// TIA Portal project "Tables" (V21)

(* hardware
DEVICE "PLC_Tables"  S7-1500 station
   slot 0: "Rail_0"  Rack  6ES7 590-1***0-0AA0
   slot 1: "PLC_Tables"  CPU 1516-3 PN/DP  6ES7 516-3AN02-0AB0  V2.9
      slot 3: "CPU display_1"  6ES7591-1BA00-0AA0
      slot 32768: "PROFINET interface_1"  X1
         slot 32769: "Port_1"  X1 P1
         slot 32770: "Port_2"  X1 P2
      slot 33024: "PROFINET interface_2"  X2
         slot 33025: "Port_1"  X2 P1
      slot 33280: "DP interface_1"  X3
      slot 34817: "Virtual CP interface port_1"  Virtual CP interface port  Virtual CP interface port
*)

// ===== PLC "PLC_Tables"  CPU 1516-3 PN/DP =====
// protected blocks, not shown: "Sealed"

VAR_GLOBAL   // PLC tag table "IO"
   "Start" AT %I0.0 : Bool;   // Start button
   "Stop" AT %I0.1 : Bool;   // Stop button, normally closed
   "DoorClosed" AT %I0.2 : Bool;   // Door switch
   "Level" AT %IW2 : Int;   // Tank level in percent
   "Motor" AT %Q0.0 : Bool;   // Motor contactor
   "Lamp" AT %Q0.1 : Bool;   // Signal lamp
   "Valve" AT %Q0.2 : Bool;   // Inlet valve
   "Fault" AT %M0.0 : Bool;   // Collected fault
   "StartEdge" AT %M0.1 : Bool;   // Edge memory of Start
   "Setpoint" AT %MW10 : Int;   // Level setpoint
   "Parts" AT %MW12 : Int;   // Parts counted
   "Speed" AT %MD20 : Real;   // Conveyor speed
   "StatusWord" AT %MW30 : Word;   // Status bits
   "Alarm" AT %M1.0 : Bool;   // Set by the sealed block
END_VAR

TYPE "RecipeStep"
   STRUCT
      target : Real;   // Speed to reach
      duration : Time;   // How long to hold it
   END_STRUCT;
END_TYPE

// folder: Common

DATA_BLOCK "LampDelay"   // DB1
{ S7_Optimized_Access := 'TRUE' }
AUTHOR : Simatic
FAMILY : IEC
NAME : IEC_TMR
VERSION : 1.0
// stored: InstanceOfName IEC_TIMER
"IEC_TIMER"
BEGIN
END_DATA_BLOCK

// folder: Data

DATA_BLOCK "Recipe"   // DB2
{ S7_Optimized_Access := 'TRUE' }
VERSION : 0.1
   VAR
      active : Bool;   // A recipe runs
      count : Int;   // Cycles run
      steps : Array[1..3] of "RecipeStep";
      limits : Struct
         low : Int;
         high : Int := 90;
      END_STRUCT;
   END_VAR
BEGIN
END_DATA_BLOCK

DATA_BLOCK "LadBoxesData"   // DB3
{ S7_Optimized_Access := 'TRUE' }
VERSION : 0.1
// stored: InstanceOfName LadBoxes
"LadBoxes"
BEGIN
END_DATA_BLOCK

// folder: (top level)

ORGANIZATION_BLOCK "Main"   // OB1, SCL, ProgramCycle
TITLE = "Main Program Sweep (Cycle)"
{ S7_Optimized_Access := 'TRUE' }
VERSION : 0.1
   VAR_INPUT
      Initial_Call : Bool;   // Initial call of this OB
      Remanence : Bool;   // =True, if remanent data are available
   END_VAR
BEGIN

    "UseRecipe"();
    "Sealed"();
    "LadBoxesData"();
    "StatusWord" := "StatusWord" OR 16#0001;
END_ORGANIZATION_BLOCK

// folder: Common

FUNCTION_BLOCK "Pulse"   // FB1, SCL
TITLE = One cycle pulse on a rising edge
{ S7_Optimized_Access := 'TRUE' }
VERSION : 0.1
   VAR_INPUT
      trigger : Bool;
   END_VAR
   VAR_OUTPUT
      q : Bool;
   END_VAR
   VAR
      last : Bool;
   END_VAR
BEGIN

    #q := #trigger AND NOT #last;
    #last := #trigger;
END_FUNCTION_BLOCK

FUNCTION "Limit" : Int   // FC1, SCL
TITLE = Clamps a value
{ S7_Optimized_Access := 'TRUE' }
VERSION : 0.1
   VAR_INPUT
      value : Int;
      low : Int;
      high : Int;
   END_VAR
BEGIN

    IF #value < #low THEN
        #Limit := #low;
    ELSIF #value > #high THEN
        #Limit := #high;
    ELSE
        #Limit := #value;
    END_IF;
END_FUNCTION

FUNCTION "Tick" : Void   // FC2, SCL
TITLE = Counts a part
{ S7_Optimized_Access := 'TRUE' }
VERSION : 0.1
BEGIN

    "Parts" := "Parts" + 1;
END_FUNCTION

// folder: Data

FUNCTION "UseRecipe" : Void   // FC3, SCL
TITLE = Runs the recipe
{ S7_Optimized_Access := 'TRUE' }
VERSION : 0.1
BEGIN

    IF "Recipe".active THEN
        "Recipe".count := "Recipe".count + 1;
        "Speed" := "Recipe".steps[1].target;
    END_IF;
    "Setpoint" := "Limit"(value := "Level", low := "Recipe".limits.low, high := "Recipe".limits.high);
END_FUNCTION

// folder: Function

FUNCTION_BLOCK "FbdLogic"   // FB13, FBD
TITLE = Function block logic
{ S7_Optimized_Access := 'TRUE' }
// Bit logic in function block diagram: gates, a set and reset box, an edge and a jump.
   VAR_INPUT
      start : Bool;
      stop : Bool;
      door : Bool;
   END_VAR
   VAR_OUTPUT
      motor : Bool;
      lamp : Bool;
      fault : Bool;
   END_VAR
   VAR
      latched : Bool;
      edgeMemory : Bool;
   END_VAR
   VAR_TEMP   // added for the SCL form of the ladder/FBD networks
      _w1 : Bool;
   END_VAR
BEGIN

REGION Network 1: Start and stop
   // OR and AND boxes drive the motor, stop negated.
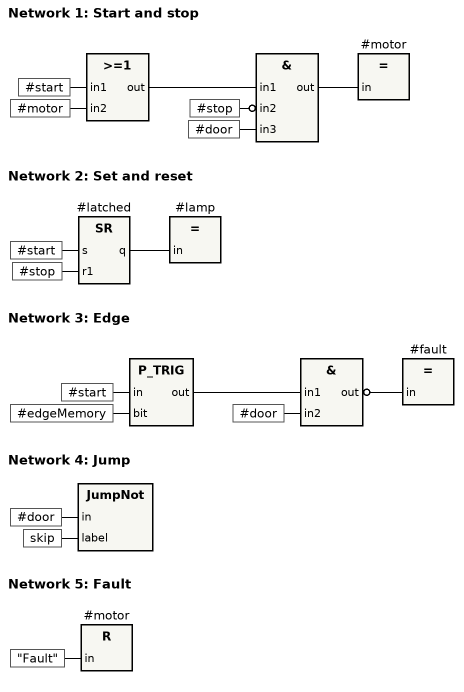
   #motor := (#start OR #motor) AND NOT #stop AND #door;
END_REGION

REGION Network 2: Set and reset
   // A set and reset box, its output on the lamp.
   IF #start THEN
       #latched := TRUE;   // SR flip-flop
   END_IF;
   IF #stop THEN #latched := FALSE; END_IF;
   #lamp := #latched;
END_REGION

REGION Network 3: Edge
   // A rising edge of start and the door, negated, is the fault.
   #_w1 := #start AND NOT #edgeMemory;   // rising edge
   #edgeMemory := #start;
   #fault := NOT (#_w1 AND #door);
END_REGION

REGION Network 4: Jump
   // Without the door closed, skip to the end.
   // no SCL statement known for JumpNot: written as a call
   JumpNot(in := #door, label := skip);
END_REGION

REGION Network 5: Fault
   // Jump target; a fault resets the motor.
   skip:
   IF "Fault" THEN #motor := FALSE; END_IF;
END_REGION
END_FUNCTION_BLOCK

FUNCTION_BLOCK "FbdBoxes"   // FB14, FBD
TITLE = Boxes
{ S7_Optimized_Access := 'TRUE' }
// Boxes in function block diagram: move, compare, add, timers, a counter and calls.
   VAR_INPUT
      level : Int;
      count : Bool;
      reset : Bool;
   END_VAR
   VAR_OUTPUT
      high : Bool;
      clamped : Int;
      done : Bool;
      pulse : Bool;
   END_VAR
   VAR
      delay : TON_TIME;
   END_VAR
   VAR RETAIN
      "counter" : CTU_INT;
   END_VAR
   VAR
      pulser : "Pulse";
      copy : Int;
      sum : Int;
   END_VAR
BEGIN

REGION Network 1: Move
   // Copies the level.
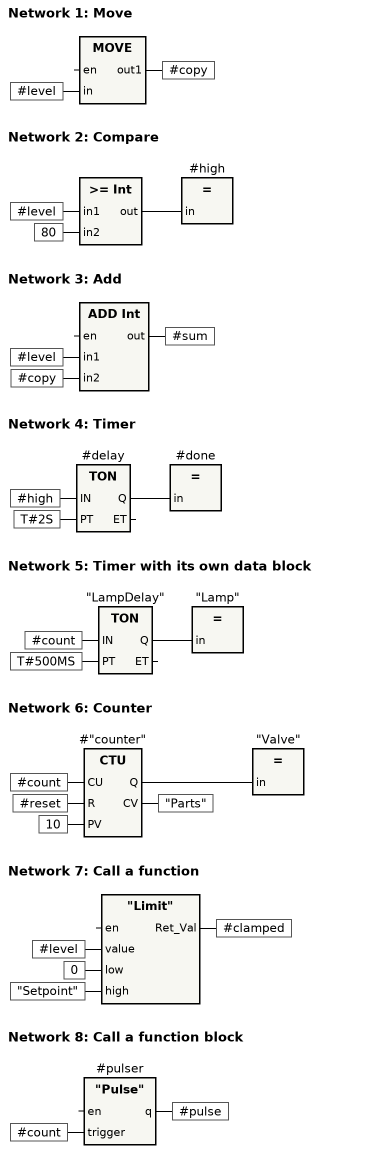
   #copy := #level;
END_REGION

REGION Network 2: Compare
   // High above 80 percent.
   #high := #level >= 80;
END_REGION

REGION Network 3: Add
   // Adds level and copy.
   #sum := #level + #copy;
END_REGION

REGION Network 4: Timer
   // Done two seconds after high, a multi-instance.
   #delay(IN := #high, PT := T#2S);   // TON
   #done := #delay.Q;
END_REGION

REGION Network 5: Timer with its own data block
   // The lamp follows count after half a second.
   "LampDelay".TON(IN := #count, PT := T#500MS);
   "Lamp" := "LampDelay".Q;
END_REGION

REGION Network 6: Counter
   // Counts parts up to ten.
   #"counter"(CU := #count, R := #reset, PV := 10, CV => "Parts");   // CTU
   "Valve" := #"counter".Q;
END_REGION

REGION Network 7: Call a function
   // Clamps the level to the setpoint.
   #clamped := "Limit"(value := #level, low := 0, high := "Setpoint");
END_REGION

REGION Network 8: Call a function block
   // A pulse on each count, a multi-instance.
   #pulser(trigger := #count, q => #pulse);   // "Pulse"
END_REGION
END_FUNCTION_BLOCK

// folder: Ladder

FUNCTION_BLOCK "LadLogic"   // FB10, LAD
TITLE = Ladder logic
{ S7_Optimized_Access := 'TRUE' }
// Bit logic in ladder: contacts, coils, an edge and a jump.
   VAR_INPUT
      start : Bool;
      stop : Bool;
      door : Bool;
   END_VAR
   VAR_OUTPUT
      motor : Bool;
      lamp : Bool;
      fault : Bool;
   END_VAR
   VAR
      latched : Bool;
      edgeMemory : Bool;
   END_VAR
   VAR_TEMP   // added for the SCL form of the ladder/FBD networks
      _w1 : Bool;
   END_VAR
BEGIN

REGION Network 1: Start and stop
   // Contacts in series and in parallel drive the motor.
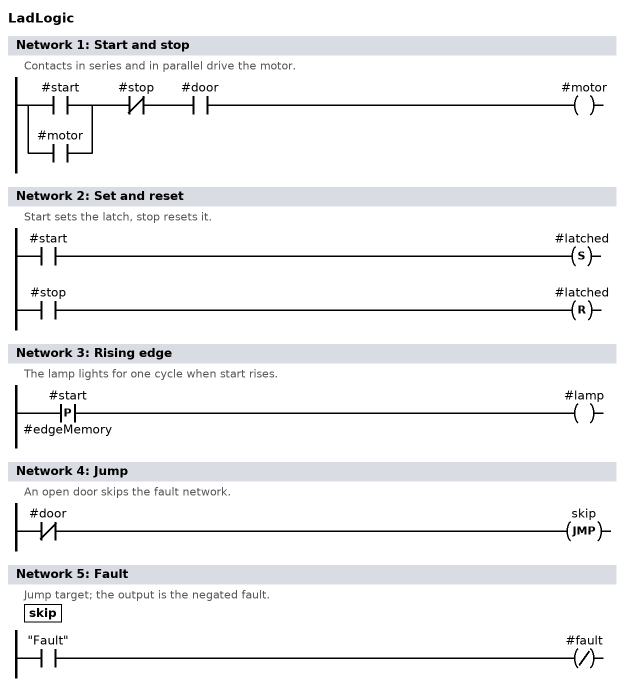
   RUNG wire#powerrail
      Contact( #start )
      wire#w1
      I_Contact( #stop )
      Contact( #door )
      Coil( #motor )
   END_RUNG
   RUNG wire#powerrail
      Contact( #motor )
   END_RUNG wire#w1
   // the same network as SCL:
   #motor := (#start OR #motor) AND NOT #stop AND #door;
END_REGION

REGION Network 2: Set and reset
   // Start sets the latch, stop resets it.
   RUNG wire#powerrail
      Contact( #start )
      S_Coil( #latched )
   END_RUNG
   RUNG wire#powerrail
      Contact( #stop )
      R_Coil( #latched )
   END_RUNG
   // the same network as SCL:
   IF #start THEN #latched := TRUE; END_IF;
   IF #stop THEN #latched := FALSE; END_IF;
END_REGION

REGION Network 3: Rising edge
   // The lamp lights for one cycle when start rises.
   RUNG wire#powerrail
      P_Contact(operand := #start, bit := #edgeMemory)
      Coil( #lamp )
   END_RUNG
   // the same network as SCL:
   #_w1 := #start AND NOT #edgeMemory;   // rising edge of #start
   #edgeMemory := #start;
   #lamp := #_w1;
END_REGION

REGION Network 4: Jump
   // An open door skips the fault network.
   RUNG wire#powerrail
      I_Contact( #door )
      JumpCoil( skip )
   END_RUNG
   // the same network as SCL:
   IF NOT #door THEN GOTO skip; END_IF;
END_REGION

REGION Network 5: Fault
   // Jump target; the output is the negated fault.
   Label( skip )
   RUNG wire#powerrail
      Contact( "Fault" )
      I_Coil( #fault )
   END_RUNG
   // the same network as SCL:
   skip:
   #fault := NOT "Fault";
END_REGION
END_FUNCTION_BLOCK

FUNCTION_BLOCK "LadBoxes"   // FB11, LAD
TITLE = Boxes
{ S7_Optimized_Access := 'TRUE' }
// Boxes in ladder: move, compare, add, timers, a counter and calls.
   VAR_INPUT
      level : Int;
      count : Bool;
      reset : Bool;
   END_VAR
   VAR_OUTPUT
      high : Bool;
      clamped : Int;
      done : Bool;
      pulse : Bool;
   END_VAR
   VAR
      delay : TON_TIME;
   END_VAR
   VAR RETAIN
      "counter" : CTU_INT;
   END_VAR
   VAR
      pulser : "Pulse";
      copy : Int;
      sum : Int;
   END_VAR
BEGIN

REGION Network 1: Move
   // Copies the level.
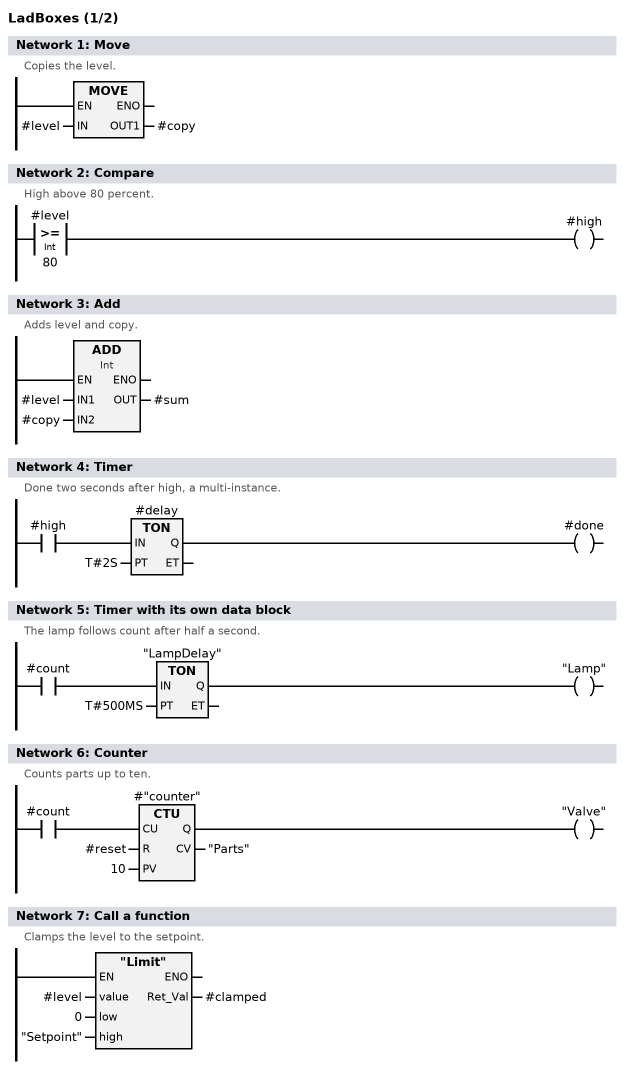
   RUNG wire#powerrail
      { S7_GenerateENO := "TRUE" } Move(in := #level, out1 => #copy)
   END_RUNG
   // the same network as SCL:
   #copy := #level;
END_REGION

REGION Network 2: Compare
   // High above 80 percent.
   RUNG wire#powerrail
      { S7_Templates := "SrcType := Int" } GE_Contact(in1 := #level, in2 := 80)
      Coil( #high )
   END_RUNG
   // the same network as SCL:
   #high := #level >= 80;
END_REGION

REGION Network 3: Add
   // Adds level and copy.
   RUNG wire#powerrail
      { S7_Templates := "SrcType := Int"; S7_GenerateENO := "TRUE" } Add(in1 := #level, in2 := #copy, out => #sum)
   END_RUNG
   // the same network as SCL:
   #sum := #level + #copy;
END_REGION

REGION Network 4: Timer
   // Done two seconds after high, a multi-instance.
   #delay(IN := #high, PT := T#2S);   // TON
   #done := #delay.Q;
END_REGION

REGION Network 5: Timer with its own data block
   // The lamp follows count after half a second.
   "LampDelay".TON(IN := #count, PT := T#500MS);
   "Lamp" := "LampDelay".Q;
END_REGION

REGION Network 6: Counter
   // Counts parts up to ten.
   #"counter"(CU := #count, R := #reset, PV := 10, CV => "Parts");   // CTU
   "Valve" := #"counter".Q;
END_REGION

REGION Network 7: Call a function
   // Clamps the level to the setpoint.
   RUNG wire#powerrail
      "Limit"(value := #level, low := 0, high := "Setpoint", Ret_Val => #clamped)
   END_RUNG
   // the same network as SCL:
   #clamped := "Limit"(value := #level, low := 0, high := "Setpoint");
END_REGION

REGION Network 8: Call a function block
   // A pulse on each count, a multi-instance.
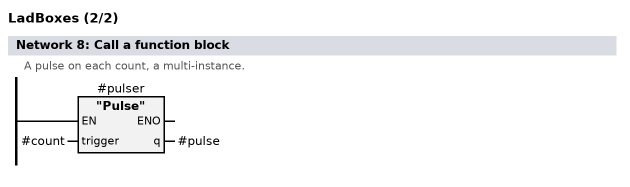
   RUNG wire#powerrail
      #pulser(trigger := #count, q => #pulse)
   END_RUNG
   // the same network as SCL:
   #pulser(trigger := #count, q => #pulse);   // "Pulse"
END_REGION
END_FUNCTION_BLOCK

FUNCTION_BLOCK "Mixed"   // FB12, LAD
TITLE = Mixed languages
{ S7_Optimized_Access := 'TRUE' }
// A ladder block with an SCL and an STL network.
   VAR_INPUT
      start : Bool;
      stop : Bool;
      door : Bool;
   END_VAR
   VAR_OUTPUT
      motor : Bool;
      lamp : Bool;
      fault : Bool;
   END_VAR
   VAR
      latched : Bool;
      edgeMemory : Bool;
   END_VAR
BEGIN

REGION Network 1: Ladder
   // A ladder network first.
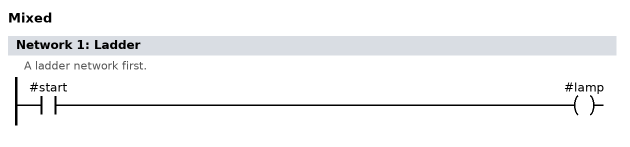
   RUNG wire#powerrail
      Contact( #start )
      Coil( #lamp )
   END_RUNG
   // the same network as SCL:
   #lamp := #start;
END_REGION

REGION Network 2 (SCL): Structured text
   // An SCL network inside a ladder block.
   #motor := #start AND NOT #stop;
END_REGION

REGION Network 3 (STL): Statement list
   // An STL network inside a ladder block.
         A     #door;
         AN    #stop;
         =     #fault;
END_REGION
END_FUNCTION_BLOCK

// folder: Sequence

FUNCTION_BLOCK "Batch"   // FB20, GRAPH_PLUS
TITLE = Batch sequence
{ S7_Optimized_Access := 'TRUE' }
// A batch sequence: fill and heat at once, mix, then drain or reject.
   VAR_INPUT
      ACK_EF : Bool := false;   // Acknowledge all errors and faults
      start : Bool;
      full : Bool;
      hot : Bool;
      quality : Bool;
      door : Bool;
      overflow : Bool;
      acknowledge : Bool;
      level : Int;
   END_VAR
   VAR_OUTPUT
      valve : Bool;
      lamp : Bool;
      heater : Bool;
      mixer : Bool;
      drain : Bool;
      alarm : Bool;
      clamped : Int;
   END_VAR
   VAR
      HMI_INFO : Array[0..10] of UInt;
      IF_PAR : G7_IfParPlus_V6;
      RT_DATA : G7_RTDataPlus_V6;   // Internal data area
      Started : G7_TransitionPlus_V6;   // Transition structure
      Ready : G7_TransitionPlus_V6;   // Transition structure
      Good : G7_TransitionPlus_V6;   // Transition structure
      Bad : G7_TransitionPlus_V6;   // Transition structure
      Empty : G7_TransitionPlus_V6;   // Transition structure
      Acknowledged : G7_TransitionPlus_V6;   // Transition structure
      Restart : G7_TransitionPlus_V6;   // Transition structure
      Idle : G7_StepPlus_V6;   // Step structure
      Fill : G7_StepPlus_V6;   // Step structure
      Heat : G7_StepPlus_V6;   // Step structure
      Mix : G7_StepPlus_V6;   // Step structure
      Discharge : G7_StepPlus_V6;   // Step structure
      Reject : G7_StepPlus_V6;   // Step structure
      Done : G7_StepPlus_V6;   // Step structure
      SINI : Array[0..3] of USInt;
      LSTT : Array[0..6] of USInt;
      ATAJ : Array[0..6] of USInt;
      ATAB : Array[0..6] of USInt;
      PSTT : Array[0..6] of USInt;
      NSTT : Array[0..6] of USInt;
      ASSJ : Array[0..6] of USInt;
      ASSB : Array[0..6] of USInt;
      PTTS : Array[0..6] of USInt;
      NTTS : Array[0..6] of USInt;
      SW_SQTS : Array[0..6] of USInt;
      SWITCH : Array[0..6] of USInt;
      TVX : Array[0..5] of USInt;
      TTX : Array[0..5] of USInt;
      TSX : Array[0..3] of USInt;
      S00X : Array[0..3] of USInt;
      SOFFX : Array[0..3] of USInt;
      SONX : Array[0..3] of USInt;
      SAX : Array[0..3] of USInt;
      SERRX : Array[0..7] of USInt;
      SMX : Array[0..7] of USInt;
      S0X : Array[0..7] of USInt;
      S1X : Array[0..7] of USInt;
      IL_ALARM_INST : Diag_Alarm;
      SUP_ALARM_INST : Diag_Alarm;
      STEP_TIME_ALARM_INST : Diag_Alarm;
      IEC_TIMER_INST : IEC_TIMER;
      TRANSACTION_FLAG : Bool := false;
   END_VAR
   // SINI[0] := 2;
   // SINI[2] := 255;
   // SINI[3] := 255;
   // LSTT[0] := 255;
   // LSTT[1] := 255;
   // LSTT[2] := 255;
   // LSTT[3] := 255;
   // LSTT[4] := 255;
   // LSTT[5] := 255;
   // ATAJ[1] := 1;
   // ATAJ[2] := 2;
   // ATAJ[3] := 3;
   // ATAJ[4] := 5;
   // ATAJ[5] := 4;
   // ATAJ[6] := 6;
   // ATAB[1] := 1;
   // ATAB[2] := 3;
   // ATAB[3] := 2;
   // ATAB[4] := 4;
   // ATAB[5] := 5;
   // ATAB[6] := 6;
   // PSTT[1] := 1;
   // PSTT[2] := 3;
   // PSTT[3] := 3;
   // PSTT[4] := 4;
   // PSTT[5] := 5;
   // PSTT[6] := 6;
   // NSTT[0] := 1;
   // NSTT[1] := 3;
   // NSTT[2] := 4;
   // NSTT[3] := 5;
   // NSTT[4] := 6;
   // NSTT[5] := 6;
   // ASSJ[1] := 2;
   // ASSJ[2] := 1;
   // ASSJ[3] := 3;
   // ASSJ[4] := 4;
   // ASSJ[5] := 5;
   // ASSJ[6] := 6;
   // ASSB[1] := 2;
   // ASSB[2] := 1;
   // ASSB[3] := 3;
   // ASSB[4] := 4;
   // ASSB[5] := 5;
   // ASSB[6] := 6;
   // PTTS[0] := 255;
   // PTTS[3] := 1;
   // PTTS[4] := 2;
   // PTTS[5] := 3;
   // PTTS[6] := 4;
   // NTTS[1] := 1;
   // NTTS[2] := 1;
   // NTTS[3] := 2;
   // NTTS[4] := 4;
   // NTTS[5] := 5;
   // NTTS[6] := 6;
   // SW_SQTS[1] := 1;
   // SW_SQTS[2] := 2;
   // SW_SQTS[3] := 3;
   // SW_SQTS[4] := 4;
   // SW_SQTS[5] := 5;
   // SW_SQTS[6] := 6;
   // SWITCH[1] := 130;
   // TVX[0] := 16#1;
   // TTX[0] := 16#1;
   // TSX[0] := 16#1;
   // S00X[0] := 16#1;
   // SOFFX[0] := 16#1;
   // SONX[0] := 16#1;
   // SAX[0] := 16#1;
   // SERRX[0] := 16#1;
   // SMX[0] := 16#1;
   // S0X[0] := 16#1;
   // S1X[0] := 16#1;
BEGIN
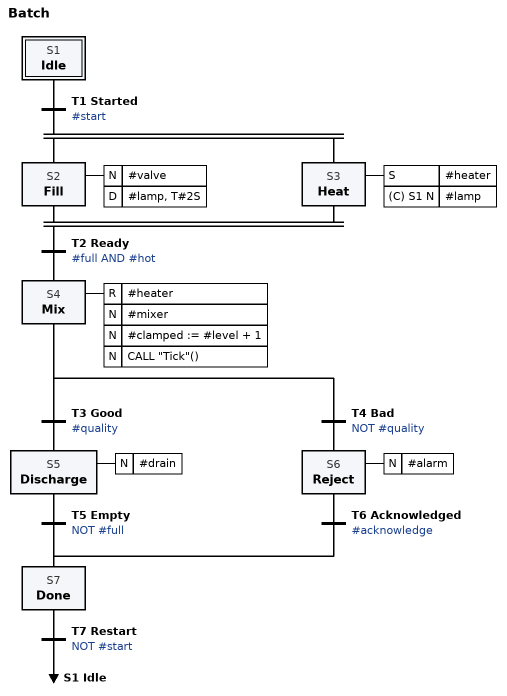
   // permanent pre-instructions
   NETWORK 1
      #lamp := #acknowledge;

   // sequencer 1
   INITIAL_STEP Idle:   // S1, max time T#10S, warning time T#7S
   END_STEP
   TRANSITION Started FROM Idle TO (Fill, Heat)   // T1
      := #start;
   END_TRANSITION
   STEP Fill:   // S2, max time T#10S, warning time T#7S
      supervision V := #overflow;
              N    #valve
              D    #lamp, T#2S
   END_STEP
   STEP Heat:   // S3, max time T#10S, warning time T#7S
      interlock C := #door;
              S    #heater
      (C) S1  N    #lamp
   END_STEP
   TRANSITION Ready FROM (Fill, Heat) TO Mix   // T2
      := #full AND #hot;
   END_TRANSITION
   STEP Mix:   // S4, max time T#10S, warning time T#7S
              R    #heater
              N    #mixer
              N    #clamped := #level + 1
              N    CALL "Tick"()
   END_STEP
   TRANSITION Good FROM Mix TO Discharge   // T3
      := #quality;
   END_TRANSITION
   TRANSITION Bad FROM Mix TO Reject   // T4
      := NOT #quality;
   END_TRANSITION
   STEP Discharge:   // S5, max time T#10S, warning time T#7S
              N    #drain
   END_STEP
   TRANSITION Empty FROM Discharge TO Done   // T5
      := NOT #full;
   END_TRANSITION
   STEP Reject:   // S6, max time T#10S, warning time T#7S
              N    #alarm
   END_STEP
   TRANSITION Acknowledged FROM Reject TO Done   // T6
      := #acknowledge;
   END_TRANSITION
   STEP Done:   // S7, max time T#10S, warning time T#7S
   END_STEP
   TRANSITION Restart FROM Done TO Idle   // T7, jump
      := NOT #start;
   END_TRANSITION

   // permanent post-instructions
   NETWORK 1
      #alarm := #overflow;
END_FUNCTION_BLOCK

// folder: Statement

FUNCTION_BLOCK "StlBasics"   // FB2, STL
TITLE = Statement list basics
{ S7_Optimized_Access := 'TRUE' }
VERSION : 0.1
// Bit logic, load and transfer, arithmetic, a jump and a call.
   VAR_INPUT
      start : Bool;
      stop : Bool;
      level : Int;
   END_VAR
   VAR_OUTPUT
      run : Bool;
      high : Bool;
      total : Int;
   END_VAR
   VAR
      count : Int;
   END_VAR
BEGIN

REGION Network 1: Latch with nesting
   // Runs from start until stop, nested in brackets.
         A(;
         O     #start;
         O     #run;
         );
         AN    #stop;
         =     #run;
END_REGION

REGION Network 2: Compare
         L     #level;
         L     80;
         >I;
         =     #high;  // above 80 percent
END_REGION

REGION Network 3: Count and transfer
         L     #count;
         L     1;
         +I;
         T     #count;
END_REGION

REGION Network 4: Jump over a call
         A     #high;
         JC    done;
         CALL  "Limit"
         ( value   := #count,
           low     := 0,
           high    := 100,
           Ret_Val := #total
         );
   done: NOP   0;
END_REGION
END_FUNCTION_BLOCK